Fanuc KAREL source: KO00024.KL

PROGRAM KO00024
%NOLOCKGROUP
VAR
  P1: XYZWPREXT
  P2: XYZWPREXT
  P3: XYZWPREXT
  P4: XYZWPREXT
  OUT: JOINTPOS
BEGIN
  OUT = FRAME(P1, P2, P3, P4)
END KO00024
